{attribute 'qualified_only'}
{attribute 'strict'}
TYPE CENTERING_ENUM :
(
	NO 	:= 0,
	TL	:= 1,
	TB	:= 2,
	ACC := 3
);
END_TYPE

(* stored: Version 1.1.0.1
   DUT CENTERING_ENUM: Id {26837bf9-1575-425e-b73b-c7c466fde73f} *)
